(* IEC 61131-3 sources: plc-vscode/tests/st/all/trust-platform/examples/OSCAT/wastewater_aeration/non-oop/src, 3 files *)

(* ---- Configuration.st ---- *)
CONFIGURATION WastewaterAerationClassicConfiguration
RESOURCE Cpu0 ON PLC
    TASK MainTask (INTERVAL := T#100ms, PRIORITY := 1);
    PROGRAM Main WITH MainTask : Main;
END_RESOURCE
END_CONFIGURATION

(* ---- Main.st ---- *)
PROGRAM Main
VAR
    OxygenDemand : HYST;
    AerationPulse : GEN_PULSE;
    DissolvedOxygen : REAL := REAL#1.5;
    BlowerCommand : BOOL;
END_VAR

OxygenDemand(In := DissolvedOxygen, HIGH_LIMIT := REAL#2.0, LOW_LIMIT := REAL#1.0);
AerationPulse(ENQ := OxygenDemand.Q, PTH := T#2s, PTL := T#3s);
BlowerCommand := AerationPulse.Q;
END_PROGRAM

(* ---- Tests.st ---- *)
TEST_PROGRAM WastewaterAerationClassicGatesPulseWithDemand
VAR
    OxygenDemand : HYST;
    AerationPulse : GEN_PULSE;
    ExpectedPulse : GEN_PULSE;
END_VAR

OxygenDemand(In := REAL#2.5, HIGH_LIMIT := REAL#2.0, LOW_LIMIT := REAL#1.0);
AerationPulse(ENQ := OxygenDemand.Q, PTH := T#2s, PTL := T#3s);
ExpectedPulse(ENQ := TRUE, PTH := T#2s, PTL := T#3s);

ASSERT_TRUE(IN := OxygenDemand.Q);
ASSERT_TRUE(IN := AerationPulse.Q = ExpectedPulse.Q);
END_TEST_PROGRAM
